FUNCTION_BLOCK FB_KUKA_REF
VAR_INPUT
	KukaToPlc			:ST_KUKATOPLC;
	PlcToKuka			:ST_PLCTOKUKA;
END_VAR
VAR_OUTPUT

END_VAR
VAR_IN_OUT

END_VAR
VAR

END_VAR

;

END_FUNCTION_BLOCK

(* stored: Version 1.1.0.1, ProductVersion 3.1.4024.15
   POU FB_KUKA_REF: Id {f45306a2-89dc-4d98-af54-e9d98824c156}, SpecialFunc None *)
